Universal Robots URScript: PrecProg.script

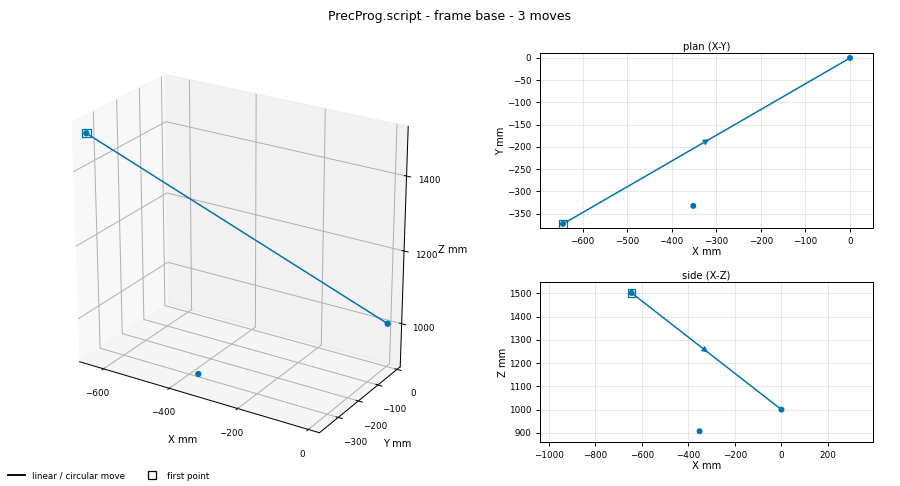
[picture p0: tool path of PrecProg.script in frame base, 3 of 6 moves have a stored position in this frame; points joined in program order, loops and branches not executed]
def PrecProg():
  # Global parameters:
  global speed_ms    = 0.250
  global speed_rads  = 0.750
  global accel_mss   = 1.200
  global accel_radss = 1.200
  global blend_radius_m = 0.001
  global ref_frame = p[0,0,0,0,0,0]

  #
  # TO REMOVE HEADER:
  # Go to "Program" -> "Post-Processor Editor"
  # Select "Universal Robots"
  # Set "INCLUDE_HEADER" to "False"
  #
  #--------------------------
  # Add any default subprograms here
  # For example, to drive a gripper as a program call:
  # def Gripper_Open():
  #   ...
  # end
  #
  # Example to drive a spray gun:
  def SprayOn(value):
    # use the value as an output:
    DO_SPRAY = 5
    if value == 0:
      set_standard_digital_out(DO_SPRAY, False)
    else:
      set_standard_digital_out(DO_SPRAY, True)
    end
  end

  # Example to drive an extruder:
  def Extruder(value):
    # use the value as an output:
    if value < 0:
      # stop extruder
    else:
      # start extruder
    end
  end

  # Example to move an external axis
  def MoveAxis(value):
    # use the value as an output:
    DO_AXIS_1 = 1
    DI_AXIS_1 = 1
    if value <= 0:
      set_standard_digital_out(DO_AXIS_1, False)

      # Wait for digital input to change state
      #while (get_standard_digital_in(DI_AXIS_1) != False):
      #  sync()
      #end
    else:
      set_standard_digital_out(DO_AXIS_1, True)

      # Wait for digital input to change state
      #while (get_standard_digital_in(DI_AXIS_1) != True):
      #  sync()
      #end
    end
  end
  #--------------------------


  # Main program:
  # Program generated by RoboDK v6.0.7 for UR10 on XX/XX/XXXX 18:00:00
  # Using nominal kinematics.
  ref_frame = p[0.000000, -0.000001, 1.000000, 1.570792, -0.005162, 0.008546]
  set_tcp(p[0.000125, -0.000375, 0.123457, -0.789761, -0.000001, 0.000002])
  movej([0.215471, -0.797247, 1.377087, -0.008727, 0.008726, 3.141593],accel_radss,speed_rads,t=0,r=0)
  movel(pose_trans(ref_frame,p[-0.640585, 0.506981, 0.371534, 0.727341, 2.187117, -0.560418]),accel_mss,speed_ms,t=0,r=0)
  movel(pose_trans(ref_frame,p[0.000500, -0.000500, 0.000250, 3.141593, 0.000137, 0.000137]),accel_mss,speed_ms,t=0,r=0.001)
  movej([-0.215468, 0.797240, -1.377065, 0.008727, -0.000002, -3.141593],accel_radss,speed_rads,t=0,r=0.001)
  movej([-0.215468, 0.797240, -1.377065, 0.008727, -0.000002, -3.141593],accel_radss,speed_rads,t=0,r=0)# end trace
  speed_ms    = 0.067
  sleep(0.002)
  sleep(1.000)
  movel(pose_trans(ref_frame,p[-0.353026, -0.090135, 0.331702, 0.124818, 2.423541, -0.239517]),accel_mss,speed_ms,t=0,r=0)
  # End of main program
end

PrecProg()
